GLOBALCONSTANTS DefaultPool_Empty_Numeric (* Numeric object pool constants (ID, Scale, Offset, Decimals) *)
  PACKAGE Uebungen::const::UT::Empty;
END_GLOBALCONSTANTS
